(* IEC 61131-3 sources: plc-st-coding-agent/progress/evidence/f14_v12_self_20261113/jobs/diagnostic_deepseek-v4pro, 15 files *)

(* ---- public-easy-01.candidate_01.st ---- *)
(* ENGINEERING_CONTRACT
Outputs by state (state is persistent across scans):
- Pump_Motor: ON in CLEANING; starts when bottleSensor TRUE from IDLE; OFF on cleaningConfirmButton. Retained while CLEANING, even if bottleSensor falls (PUB001/PUB002).
- Filling_Valve: ON in FILLING; starts on cleaningConfirmButton in CLEANING; OFF on fillingConfirmButton (PUB002/PUB003).
- Capping_Machine: ON in CAPPING; starts on fillingConfirmButton in FILLING; OFF on cappingConfirmButton (PUB003/PUB004).
- Packing_Machine: ON in PACKING; starts on cappingConfirmButton in CAPPING; OFF on packingConfirmButton (PUB004/PUB005).
- Completion_Light: ON in COMPLETE; starts on packingConfirmButton in PACKING; reset by finishedButton (PUB005/PUB006/PUB007).
Same-scan priority: one state transition per call via ELSIF chain; outputs are assigned after transition using final state.
Buttons are treated as level-sensitive; pulse width/protocol unspecified.
*)
(* CONTRACT_RULES [] *)

FUNCTION_BLOCK FillingLineControl
VAR_INPUT
    bottleSensor: BOOL;
    cleaningConfirmButton: BOOL;
    fillingConfirmButton: BOOL;
    cappingConfirmButton: BOOL;
    packingConfirmButton: BOOL;
    finishedButton: BOOL;
END_VAR
VAR_OUTPUT
    Pump_Motor: BOOL;
    Filling_Valve: BOOL;
    Capping_Machine: BOOL;
    Packing_Machine: BOOL;
    Completion_Light: BOOL;
END_VAR
VAR
    step: INT := 0; (* 0=IDLE, 1=CLEANING, 2=FILLING, 3=CAPPING, 4=PACKING, 5=COMPLETE *)
    bottleTrig: R_TRIG;
END_VAR

(* State transitions: at most one per scan *)
bottleTrig(CLK := bottleSensor);

IF step = 0 THEN
    IF bottleTrig.Q THEN
        step := 1;
    END_IF;
ELSIF step = 1 THEN
    IF cleaningConfirmButton THEN
        step := 2;
    END_IF;
ELSIF step = 2 THEN
    IF fillingConfirmButton THEN
        step := 3;
    END_IF;
ELSIF step = 3 THEN
    IF cappingConfirmButton THEN
        step := 4;
    END_IF;
ELSIF step = 4 THEN
    IF packingConfirmButton THEN
        step := 5;
    END_IF;
ELSIF step = 5 THEN
    IF finishedButton THEN
        step := 0;
    END_IF;
END_IF;

(* Output mapping based on final state *)
CASE step OF
    0:
        Pump_Motor := FALSE;
        Filling_Valve := FALSE;
        Capping_Machine := FALSE;
        Packing_Machine := FALSE;
        Completion_Light := FALSE;

    1:
        Pump_Motor := TRUE;
        Filling_Valve := FALSE;
        Capping_Machine := FALSE;
        Packing_Machine := FALSE;
        Completion_Light := FALSE;

    2:
        Pump_Motor := FALSE;
        Filling_Valve := TRUE;
        Capping_Machine := FALSE;
        Packing_Machine := FALSE;
        Completion_Light := FALSE;

    3:
        Pump_Motor := FALSE;
        Filling_Valve := FALSE;
        Capping_Machine := TRUE;
        Packing_Machine := FALSE;
        Completion_Light := FALSE;

    4:
        Pump_Motor := FALSE;
        Filling_Valve := FALSE;
        Capping_Machine := FALSE;
        Packing_Machine := TRUE;
        Completion_Light := FALSE;

    5:
        Pump_Motor := FALSE;
        Filling_Valve := FALSE;
        Capping_Machine := FALSE;
        Packing_Machine := FALSE;
        Completion_Light := TRUE;

    ELSE
        Pump_Motor := FALSE;
        Filling_Valve := FALSE;
        Capping_Machine := FALSE;
        Packing_Machine := FALSE;
        Completion_Light := FALSE;
END_CASE;

END_FUNCTION_BLOCK

(* ---- public-easy-01.candidate_02.st ---- *)
(* ENGINEERING_CONTRACT
Outputs by state (state is persistent across scans):
- Pump_Motor: ON in CLEANING; starts when bottleSensor TRUE from IDLE; OFF on cleaningConfirmButton. Retained while CLEANING, even if bottleSensor falls (PUB001/PUB002).
- Filling_Valve: ON in FILLING; starts on cleaningConfirmButton in CLEANING; OFF on fillingConfirmButton (PUB002/PUB003).
- Capping_Machine: ON in CAPPING; starts on fillingConfirmButton in FILLING; OFF on cappingConfirmButton (PUB003/PUB004).
- Packing_Machine: ON in PACKING; starts on cappingConfirmButton in CAPPING; OFF on packingConfirmButton (PUB004/PUB005).
- Completion_Light: ON in COMPLETE; starts on packingConfirmButton in PACKING; reset by finishedButton (PUB005/PUB006/PUB007).
Same-scan priority: one state transition per call via ELSIF chain; outputs are assigned after transition using final state.
Buttons are treated as level-sensitive; pulse width/protocol unspecified.
*)
(* CONTRACT_RULES [] *)

FUNCTION_BLOCK FillingLineControl
VAR_INPUT
    bottleSensor: BOOL;
    cleaningConfirmButton: BOOL;
    fillingConfirmButton: BOOL;
    cappingConfirmButton: BOOL;
    packingConfirmButton: BOOL;
    finishedButton: BOOL;
END_VAR
VAR_OUTPUT
    Pump_Motor: BOOL;
    Filling_Valve: BOOL;
    Capping_Machine: BOOL;
    Packing_Machine: BOOL;
    Completion_Light: BOOL;
END_VAR
VAR
    step: INT := 0; (* 0=IDLE, 1=CLEANING, 2=FILLING, 3=CAPPING, 4=PACKING, 5=COMPLETE *)
END_VAR

(* State transitions: at most one per scan *)
IF step = 0 THEN
    IF bottleSensor THEN
        step := 1;
    END_IF;
ELSIF step = 1 THEN
    IF cleaningConfirmButton THEN
        step := 2;
    END_IF;
ELSIF step = 2 THEN
    IF fillingConfirmButton THEN
        step := 3;
    END_IF;
ELSIF step = 3 THEN
    IF cappingConfirmButton THEN
        step := 4;
    END_IF;
ELSIF step = 4 THEN
    IF packingConfirmButton THEN
        step := 5;
    END_IF;
ELSIF step = 5 THEN
    IF finishedButton THEN
        step := 0;
    END_IF;
END_IF;

(* Output mapping based on final state *)
CASE step OF
    0:
        Pump_Motor := FALSE;
        Filling_Valve := FALSE;
        Capping_Machine := FALSE;
        Packing_Machine := FALSE;
        Completion_Light := FALSE;

    1:
        Pump_Motor := TRUE;
        Filling_Valve := FALSE;
        Capping_Machine := FALSE;
        Packing_Machine := FALSE;
        Completion_Light := FALSE;

    2:
        Pump_Motor := FALSE;
        Filling_Valve := TRUE;
        Capping_Machine := FALSE;
        Packing_Machine := FALSE;
        Completion_Light := FALSE;

    3:
        Pump_Motor := FALSE;
        Filling_Valve := FALSE;
        Capping_Machine := TRUE;
        Packing_Machine := FALSE;
        Completion_Light := FALSE;

    4:
        Pump_Motor := FALSE;
        Filling_Valve := FALSE;
        Capping_Machine := FALSE;
        Packing_Machine := TRUE;
        Completion_Light := FALSE;

    5:
        Pump_Motor := FALSE;
        Filling_Valve := FALSE;
        Capping_Machine := FALSE;
        Packing_Machine := FALSE;
        Completion_Light := TRUE;

    ELSE
        Pump_Motor := FALSE;
        Filling_Valve := FALSE;
        Capping_Machine := FALSE;
        Packing_Machine := FALSE;
        Completion_Light := FALSE;
END_CASE;

END_FUNCTION_BLOCK

(* ---- public-easy-01.candidate_03.st ---- *)
(* ENGINEERING_CONTRACT
Outputs by state (state is persistent across scans):
- Pump_Motor: ON in CLEANING; starts when bottleSensor TRUE from IDLE; OFF on cleaningConfirmButton. Retained while CLEANING, even if bottleSensor falls (PUB001/PUB002).
- Filling_Valve: ON in FILLING; starts on cleaningConfirmButton in CLEANING; OFF on fillingConfirmButton (PUB002/PUB003).
- Capping_Machine: ON in CAPPING; starts on fillingConfirmButton in FILLING; OFF on cappingConfirmButton (PUB003/PUB004).
- Packing_Machine: ON in PACKING; starts on cappingConfirmButton in CAPPING; OFF on packingConfirmButton (PUB004/PUB005).
- Completion_Light: ON in COMPLETE; starts on packingConfirmButton in PACKING; reset by finishedButton (PUB005/PUB006/PUB007).
Same-scan priority: one state transition per call via ELSIF chain; outputs are assigned after transition using final state.
Buttons are treated as level-sensitive; pulse width/protocol unspecified.
*)
(* CONTRACT_RULES [] *)

FUNCTION_BLOCK FillingLineControl
VAR_INPUT
    bottleSensor: BOOL;
    cleaningConfirmButton: BOOL;
    fillingConfirmButton: BOOL;
    cappingConfirmButton: BOOL;
    packingConfirmButton: BOOL;
    finishedButton: BOOL;
END_VAR
VAR_OUTPUT
    Pump_Motor: BOOL;
    Filling_Valve: BOOL;
    Capping_Machine: BOOL;
    Packing_Machine: BOOL;
    Completion_Light: BOOL;
END_VAR
VAR
    step: INT := 0; (* 0=IDLE, 1=CLEANING, 2=FILLING, 3=CAPPING, 4=PACKING, 5=COMPLETE *)
    local_i: INT;
END_VAR

(* State transitions: at most one per scan *)
FOR local_i := 0 TO 5 DO
    IF step = 0 THEN
        IF bottleSensor THEN
            step := 1;
        END_IF;
    ELSIF step = 1 THEN
        IF cleaningConfirmButton THEN
            step := 2;
        END_IF;
    ELSIF step = 2 THEN
        IF fillingConfirmButton THEN
            step := 3;
        END_IF;
    ELSIF step = 3 THEN
        IF cappingConfirmButton THEN
            step := 4;
        END_IF;
    ELSIF step = 4 THEN
        IF packingConfirmButton THEN
            step := 5;
        END_IF;
    ELSIF step = 5 THEN
        IF finishedButton THEN
            step := 0;
        END_IF;
    END_IF;
END_FOR;

(* Output mapping based on final state *)
CASE step OF
    0:
        Pump_Motor := FALSE;
        Filling_Valve := FALSE;
        Capping_Machine := FALSE;
        Packing_Machine := FALSE;
        Completion_Light := FALSE;

    1:
        Pump_Motor := TRUE;
        Filling_Valve := FALSE;
        Capping_Machine := FALSE;
        Packing_Machine := FALSE;
        Completion_Light := FALSE;

    2:
        Pump_Motor := FALSE;
        Filling_Valve := TRUE;
        Capping_Machine := FALSE;
        Packing_Machine := FALSE;
        Completion_Light := FALSE;

    3:
        Pump_Motor := FALSE;
        Filling_Valve := FALSE;
        Capping_Machine := TRUE;
        Packing_Machine := FALSE;
        Completion_Light := FALSE;

    4:
        Pump_Motor := FALSE;
        Filling_Valve := FALSE;
        Capping_Machine := FALSE;
        Packing_Machine := TRUE;
        Completion_Light := FALSE;

    5:
        Pump_Motor := FALSE;
        Filling_Valve := FALSE;
        Capping_Machine := FALSE;
        Packing_Machine := FALSE;
        Completion_Light := TRUE;

    ELSE
        Pump_Motor := FALSE;
        Filling_Valve := FALSE;
        Capping_Machine := FALSE;
        Packing_Machine := FALSE;
        Completion_Light := FALSE;
END_CASE;

END_FUNCTION_BLOCK

(* ---- public-easy-01.patch_base_01.st ---- *)
(* ENGINEERING_CONTRACT
Outputs by state (state is persistent across scans):
- Pump_Motor: ON in CLEANING; starts when bottleSensor TRUE from IDLE; OFF on cleaningConfirmButton. Retained while CLEANING, even if bottleSensor falls (PUB001/PUB002).
- Filling_Valve: ON in FILLING; starts on cleaningConfirmButton in CLEANING; OFF on fillingConfirmButton (PUB002/PUB003).
- Capping_Machine: ON in CAPPING; starts on fillingConfirmButton in FILLING; OFF on cappingConfirmButton (PUB003/PUB004).
- Packing_Machine: ON in PACKING; starts on cappingConfirmButton in CAPPING; OFF on packingConfirmButton (PUB004/PUB005).
- Completion_Light: ON in COMPLETE; starts on packingConfirmButton in PACKING; reset by finishedButton (PUB005/PUB006/PUB007).
Same-scan priority: one state transition per call via ELSIF chain; outputs are assigned after transition using final state.
Buttons are treated as level-sensitive; pulse width/protocol unspecified.
*)
(* CONTRACT_RULES [] *)

FUNCTION_BLOCK FillingLineControl
VAR_INPUT
    bottleSensor: BOOL;
    cleaningConfirmButton: BOOL;
    fillingConfirmButton: BOOL;
    cappingConfirmButton: BOOL;
    packingConfirmButton: BOOL;
    finishedButton: BOOL;
END_VAR
VAR_OUTPUT
    Pump_Motor: BOOL;
    Filling_Valve: BOOL;
    Capping_Machine: BOOL;
    Packing_Machine: BOOL;
    Completion_Light: BOOL;
END_VAR
VAR
    step: INT := 0; (* 0=IDLE, 1=CLEANING, 2=FILLING, 3=CAPPING, 4=PACKING, 5=COMPLETE *)
END_VAR

(* State transitions: at most one per scan *)
IF step = 0 THEN
    IF bottleSensor THEN
        step := 1;
    END_IF;
ELSIF step = 1 THEN
    IF cleaningConfirmButton THEN
        step := 2;
    END_IF;
ELSIF step = 2 THEN
    IF fillingConfirmButton THEN
        step := 3;
    END_IF;
ELSIF step = 3 THEN
    IF cappingConfirmButton THEN
        step := 4;
    END_IF;
ELSIF step = 4 THEN
    IF packingConfirmButton THEN
        step := 5;
    END_IF;
ELSIF step = 5 THEN
    IF finishedButton THEN
        step := 0;
    END_IF;
END_IF;

(* Output mapping based on final state *)
CASE step OF
    0:
        Pump_Motor := FALSE;
        Filling_Valve := FALSE;
        Capping_Machine := FALSE;
        Packing_Machine := FALSE;
        Completion_Light := FALSE;

    1:
        Pump_Motor := TRUE;
        Filling_Valve := FALSE;
        Capping_Machine := FALSE;
        Packing_Machine := FALSE;
        Completion_Light := FALSE;

    2:
        Pump_Motor := FALSE;
        Filling_Valve := TRUE;
        Capping_Machine := FALSE;
        Packing_Machine := FALSE;
        Completion_Light := FALSE;

    3:
        Pump_Motor := FALSE;
        Filling_Valve := FALSE;
        Capping_Machine := TRUE;
        Packing_Machine := FALSE;
        Completion_Light := FALSE;

    4:
        Pump_Motor := FALSE;
        Filling_Valve := FALSE;
        Capping_Machine := FALSE;
        Packing_Machine := TRUE;
        Completion_Light := FALSE;

    5:
        Pump_Motor := FALSE;
        Filling_Valve := FALSE;
        Capping_Machine := FALSE;
        Packing_Machine := FALSE;
        Completion_Light := TRUE;

    ELSE
        Pump_Motor := FALSE;
        Filling_Valve := FALSE;
        Capping_Machine := FALSE;
        Packing_Machine := FALSE;
        Completion_Light := FALSE;
END_CASE;

END_FUNCTION_BLOCK

(* ---- public-easy-01.patch_base_02.st ---- *)
(* ENGINEERING_CONTRACT
Outputs by state (state is persistent across scans):
- Pump_Motor: ON in CLEANING; starts when bottleSensor TRUE from IDLE; OFF on cleaningConfirmButton. Retained while CLEANING, even if bottleSensor falls (PUB001/PUB002).
- Filling_Valve: ON in FILLING; starts on cleaningConfirmButton in CLEANING; OFF on fillingConfirmButton (PUB002/PUB003).
- Capping_Machine: ON in CAPPING; starts on fillingConfirmButton in FILLING; OFF on cappingConfirmButton (PUB003/PUB004).
- Packing_Machine: ON in PACKING; starts on cappingConfirmButton in CAPPING; OFF on packingConfirmButton (PUB004/PUB005).
- Completion_Light: ON in COMPLETE; starts on packingConfirmButton in PACKING; reset by finishedButton (PUB005/PUB006/PUB007).
Same-scan priority: one state transition per call via ELSIF chain; outputs are assigned after transition using final state.
Buttons are treated as level-sensitive; pulse width/protocol unspecified.
*)
(* CONTRACT_RULES [] *)

FUNCTION_BLOCK FillingLineControl
VAR_INPUT
    bottleSensor: BOOL;
    cleaningConfirmButton: BOOL;
    fillingConfirmButton: BOOL;
    cappingConfirmButton: BOOL;
    packingConfirmButton: BOOL;
    finishedButton: BOOL;
END_VAR
VAR_OUTPUT
    Pump_Motor: BOOL;
    Filling_Valve: BOOL;
    Capping_Machine: BOOL;
    Packing_Machine: BOOL;
    Completion_Light: BOOL;
END_VAR
VAR
    step: INT := 0; (* 0=IDLE, 1=CLEANING, 2=FILLING, 3=CAPPING, 4=PACKING, 5=COMPLETE *)
    bottleTrig: R_TRIG;
END_VAR

(* State transitions: at most one per scan *)
bottleTrig(CLK := bottleSensor);

IF step = 0 THEN
    IF bottleTrig.Q THEN
        step := 1;
    END_IF;
ELSIF step = 1 THEN
    IF cleaningConfirmButton THEN
        step := 2;
    END_IF;
ELSIF step = 2 THEN
    IF fillingConfirmButton THEN
        step := 3;
    END_IF;
ELSIF step = 3 THEN
    IF cappingConfirmButton THEN
        step := 4;
    END_IF;
ELSIF step = 4 THEN
    IF packingConfirmButton THEN
        step := 5;
    END_IF;
ELSIF step = 5 THEN
    IF finishedButton THEN
        step := 0;
    END_IF;
END_IF;

(* Output mapping based on final state *)
CASE step OF
    0:
        Pump_Motor := FALSE;
        Filling_Valve := FALSE;
        Capping_Machine := FALSE;
        Packing_Machine := FALSE;
        Completion_Light := FALSE;

    1:
        Pump_Motor := TRUE;
        Filling_Valve := FALSE;
        Capping_Machine := FALSE;
        Packing_Machine := FALSE;
        Completion_Light := FALSE;

    2:
        Pump_Motor := FALSE;
        Filling_Valve := TRUE;
        Capping_Machine := FALSE;
        Packing_Machine := FALSE;
        Completion_Light := FALSE;

    3:
        Pump_Motor := FALSE;
        Filling_Valve := FALSE;
        Capping_Machine := TRUE;
        Packing_Machine := FALSE;
        Completion_Light := FALSE;

    4:
        Pump_Motor := FALSE;
        Filling_Valve := FALSE;
        Capping_Machine := FALSE;
        Packing_Machine := TRUE;
        Completion_Light := FALSE;

    5:
        Pump_Motor := FALSE;
        Filling_Valve := FALSE;
        Capping_Machine := FALSE;
        Packing_Machine := FALSE;
        Completion_Light := TRUE;

    ELSE
        Pump_Motor := FALSE;
        Filling_Valve := FALSE;
        Capping_Machine := FALSE;
        Packing_Machine := FALSE;
        Completion_Light := FALSE;
END_CASE;

END_FUNCTION_BLOCK

(* ---- public-easy-01.patch_base_03.st ---- *)
(* ENGINEERING_CONTRACT
Outputs by state (state is persistent across scans):
- Pump_Motor: ON in CLEANING; starts when bottleSensor TRUE from IDLE; OFF on cleaningConfirmButton. Retained while CLEANING, even if bottleSensor falls (PUB001/PUB002).
- Filling_Valve: ON in FILLING; starts on cleaningConfirmButton in CLEANING; OFF on fillingConfirmButton (PUB002/PUB003).
- Capping_Machine: ON in CAPPING; starts on fillingConfirmButton in FILLING; OFF on cappingConfirmButton (PUB003/PUB004).
- Packing_Machine: ON in PACKING; starts on cappingConfirmButton in CAPPING; OFF on packingConfirmButton (PUB004/PUB005).
- Completion_Light: ON in COMPLETE; starts on packingConfirmButton in PACKING; reset by finishedButton (PUB005/PUB006/PUB007).
Same-scan priority: one state transition per call via ELSIF chain; outputs are assigned after transition using final state.
Buttons are treated as level-sensitive; pulse width/protocol unspecified.
*)
(* CONTRACT_RULES [] *)

FUNCTION_BLOCK FillingLineControl
VAR_INPUT
    bottleSensor: BOOL;
    cleaningConfirmButton: BOOL;
    fillingConfirmButton: BOOL;
    cappingConfirmButton: BOOL;
    packingConfirmButton: BOOL;
    finishedButton: BOOL;
END_VAR
VAR_OUTPUT
    Pump_Motor: BOOL;
    Filling_Valve: BOOL;
    Capping_Machine: BOOL;
    Packing_Machine: BOOL;
    Completion_Light: BOOL;
END_VAR
VAR
    step: INT := 0; (* 0=IDLE, 1=CLEANING, 2=FILLING, 3=CAPPING, 4=PACKING, 5=COMPLETE *)
END_VAR

(* State transitions: at most one per scan *)
IF step = 0 THEN
    IF bottleSensor THEN
        step := 1;
    END_IF;
ELSIF step = 1 THEN
    IF cleaningConfirmButton THEN
        step := 2;
    END_IF;
ELSIF step = 2 THEN
    IF fillingConfirmButton THEN
        step := 3;
    END_IF;
ELSIF step = 3 THEN
    IF cappingConfirmButton THEN
        step := 4;
    END_IF;
ELSIF step = 4 THEN
    IF packingConfirmButton THEN
        step := 5;
    END_IF;
ELSIF step = 5 THEN
    IF finishedButton THEN
        step := 0;
    END_IF;
END_IF;

(* Output mapping based on final state *)
CASE step OF
    0:
        Pump_Motor := FALSE;
        Filling_Valve := FALSE;
        Capping_Machine := FALSE;
        Packing_Machine := FALSE;
        Completion_Light := FALSE;

    1:
        Pump_Motor := TRUE;
        Filling_Valve := FALSE;
        Capping_Machine := FALSE;
        Packing_Machine := FALSE;
        Completion_Light := FALSE;

    2:
        Pump_Motor := FALSE;
        Filling_Valve := TRUE;
        Capping_Machine := FALSE;
        Packing_Machine := FALSE;
        Completion_Light := FALSE;

    3:
        Pump_Motor := FALSE;
        Filling_Valve := FALSE;
        Capping_Machine := TRUE;
        Packing_Machine := FALSE;
        Completion_Light := FALSE;

    4:
        Pump_Motor := FALSE;
        Filling_Valve := FALSE;
        Capping_Machine := FALSE;
        Packing_Machine := TRUE;
        Completion_Light := FALSE;

    5:
        Pump_Motor := FALSE;
        Filling_Valve := FALSE;
        Capping_Machine := FALSE;
        Packing_Machine := FALSE;
        Completion_Light := TRUE;

    ELSE
        Pump_Motor := FALSE;
        Filling_Valve := FALSE;
        Capping_Machine := FALSE;
        Packing_Machine := FALSE;
        Completion_Light := FALSE;
END_CASE;

END_FUNCTION_BLOCK

(* ---- public-easy-01.raw_candidate_01.st ---- *)
(* ENGINEERING_CONTRACT
Outputs by state (state is persistent across scans):
- Pump_Motor: ON in CLEANING; starts when bottleSensor TRUE from IDLE; OFF on cleaningConfirmButton. Retained while CLEANING, even if bottleSensor falls (PUB001/PUB002).
- Filling_Valve: ON in FILLING; starts on cleaningConfirmButton in CLEANING; OFF on fillingConfirmButton (PUB002/PUB003).
- Capping_Machine: ON in CAPPING; starts on fillingConfirmButton in FILLING; OFF on cappingConfirmButton (PUB003/PUB004).
- Packing_Machine: ON in PACKING; starts on cappingConfirmButton in CAPPING; OFF on packingConfirmButton (PUB004/PUB005).
- Completion_Light: ON in COMPLETE; starts on packingConfirmButton in PACKING; reset by finishedButton (PUB005/PUB006/PUB007).
Same-scan priority: one state transition per call via ELSIF chain; outputs are assigned after transition using final state.
Buttons are treated as level-sensitive; pulse width/protocol unspecified.
*)
(* CONTRACT_RULES [] *)

FUNCTION_BLOCK FillingLineControl
VAR_INPUT
    bottleSensor: BOOL;
    cleaningConfirmButton: BOOL;
    fillingConfirmButton: BOOL;
    cappingConfirmButton: BOOL;
    packingConfirmButton: BOOL;
    finishedButton: BOOL;
END_VAR
VAR_OUTPUT
    Pump_Motor: BOOL;
    Filling_Valve: BOOL;
    Capping_Machine: BOOL;
    Packing_Machine: BOOL;
    Completion_Light: BOOL;
END_VAR
VAR
    step: INT := 0; (* 0=IDLE, 1=CLEANING, 2=FILLING, 3=CAPPING, 4=PACKING, 5=COMPLETE *)
    bottleTrig: R_TRIG;
END_VAR

(* State transitions: at most one per scan *)
bottleTrig(CLK := bottleSensor);

IF step = 0 THEN
    IF bottleTrig.Q THEN
        step := 1;
    END_IF;
ELSIF step = 1 THEN
    IF cleaningConfirmButton THEN
        step := 2;
    END_IF;
ELSIF step = 2 THEN
    IF fillingConfirmButton THEN
        step := 3;
    END_IF;
ELSIF step = 3 THEN
    IF cappingConfirmButton THEN
        step := 4;
    END_IF;
ELSIF step = 4 THEN
    IF packingConfirmButton THEN
        step := 5;
    END_IF;
ELSIF step = 5 THEN
    IF finishedButton THEN
        step := 0;
    END_IF;
END_IF;

(* Output mapping based on final state *)
CASE step OF
    0:
        Pump_Motor := FALSE;
        Filling_Valve := FALSE;
        Capping_Machine := FALSE;
        Packing_Machine := FALSE;
        Completion_Light := FALSE;

    1:
        Pump_Motor := TRUE;
        Filling_Valve := FALSE;
        Capping_Machine := FALSE;
        Packing_Machine := FALSE;
        Completion_Light := FALSE;

    2:
        Pump_Motor := FALSE;
        Filling_Valve := TRUE;
        Capping_Machine := FALSE;
        Packing_Machine := FALSE;
        Completion_Light := FALSE;

    3:
        Pump_Motor := FALSE;
        Filling_Valve := FALSE;
        Capping_Machine := TRUE;
        Packing_Machine := FALSE;
        Completion_Light := FALSE;

    4:
        Pump_Motor := FALSE;
        Filling_Valve := FALSE;
        Capping_Machine := FALSE;
        Packing_Machine := TRUE;
        Completion_Light := FALSE;

    5:
        Pump_Motor := FALSE;
        Filling_Valve := FALSE;
        Capping_Machine := FALSE;
        Packing_Machine := FALSE;
        Completion_Light := TRUE;

    ELSE
        Pump_Motor := FALSE;
        Filling_Valve := FALSE;
        Capping_Machine := FALSE;
        Packing_Machine := FALSE;
        Completion_Light := FALSE;
END_CASE;

END_FUNCTION_BLOCK

(* ---- public-easy-01.raw_candidate_02.st ---- *)
(* ENGINEERING_CONTRACT
Outputs by state (state is persistent across scans):
- Pump_Motor: ON in CLEANING; starts when bottleSensor TRUE from IDLE; OFF on cleaningConfirmButton. Retained while CLEANING, even if bottleSensor falls (PUB001/PUB002).
- Filling_Valve: ON in FILLING; starts on cleaningConfirmButton in CLEANING; OFF on fillingConfirmButton (PUB002/PUB003).
- Capping_Machine: ON in CAPPING; starts on fillingConfirmButton in FILLING; OFF on cappingConfirmButton (PUB003/PUB004).
- Packing_Machine: ON in PACKING; starts on cappingConfirmButton in CAPPING; OFF on packingConfirmButton (PUB004/PUB005).
- Completion_Light: ON in COMPLETE; starts on packingConfirmButton in PACKING; reset by finishedButton (PUB005/PUB006/PUB007).
Same-scan priority: one state transition per call via ELSIF chain; outputs are assigned after transition using final state.
Buttons are treated as level-sensitive; pulse width/protocol unspecified.
*)
(* CONTRACT_RULES [] *)

FUNCTION_BLOCK FillingLineControl
VAR_INPUT
    bottleSensor: BOOL;
    cleaningConfirmButton: BOOL;
    fillingConfirmButton: BOOL;
    cappingConfirmButton: BOOL;
    packingConfirmButton: BOOL;
    finishedButton: BOOL;
END_VAR
VAR_OUTPUT
    Pump_Motor: BOOL;
    Filling_Valve: BOOL;
    Capping_Machine: BOOL;
    Packing_Machine: BOOL;
    Completion_Light: BOOL;
END_VAR
VAR
    step: INT := 0; (* 0=IDLE, 1=CLEANING, 2=FILLING, 3=CAPPING, 4=PACKING, 5=COMPLETE *)
END_VAR

(* State transitions: at most one per scan *)
IF step = 0 THEN
    IF bottleSensor THEN
        step := 1;
    END_IF;
ELSIF step = 1 THEN
    IF cleaningConfirmButton THEN
        step := 2;
    END_IF;
ELSIF step = 2 THEN
    IF fillingConfirmButton THEN
        step := 3;
    END_IF;
ELSIF step = 3 THEN
    IF cappingConfirmButton THEN
        step := 4;
    END_IF;
ELSIF step = 4 THEN
    IF packingConfirmButton THEN
        step := 5;
    END_IF;
ELSIF step = 5 THEN
    IF finishedButton THEN
        step := 0;
    END_IF;
END_IF;

(* Output mapping based on final state *)
CASE step OF
    0:
        Pump_Motor := FALSE;
        Filling_Valve := FALSE;
        Capping_Machine := FALSE;
        Packing_Machine := FALSE;
        Completion_Light := FALSE;

    1:
        Pump_Motor := TRUE;
        Filling_Valve := FALSE;
        Capping_Machine := FALSE;
        Packing_Machine := FALSE;
        Completion_Light := FALSE;

    2:
        Pump_Motor := FALSE;
        Filling_Valve := TRUE;
        Capping_Machine := FALSE;
        Packing_Machine := FALSE;
        Completion_Light := FALSE;

    3:
        Pump_Motor := FALSE;
        Filling_Valve := FALSE;
        Capping_Machine := TRUE;
        Packing_Machine := FALSE;
        Completion_Light := FALSE;

    4:
        Pump_Motor := FALSE;
        Filling_Valve := FALSE;
        Capping_Machine := FALSE;
        Packing_Machine := TRUE;
        Completion_Light := FALSE;

    5:
        Pump_Motor := FALSE;
        Filling_Valve := FALSE;
        Capping_Machine := FALSE;
        Packing_Machine := FALSE;
        Completion_Light := TRUE;

    ELSE
        Pump_Motor := FALSE;
        Filling_Valve := FALSE;
        Capping_Machine := FALSE;
        Packing_Machine := FALSE;
        Completion_Light := FALSE;
END_CASE;

END_FUNCTION_BLOCK

(* ---- public-easy-01.raw_candidate_03.st ---- *)
(* ENGINEERING_CONTRACT
Outputs by state (state is persistent across scans):
- Pump_Motor: ON in CLEANING; starts when bottleSensor TRUE from IDLE; OFF on cleaningConfirmButton. Retained while CLEANING, even if bottleSensor falls (PUB001/PUB002).
- Filling_Valve: ON in FILLING; starts on cleaningConfirmButton in CLEANING; OFF on fillingConfirmButton (PUB002/PUB003).
- Capping_Machine: ON in CAPPING; starts on fillingConfirmButton in FILLING; OFF on cappingConfirmButton (PUB003/PUB004).
- Packing_Machine: ON in PACKING; starts on cappingConfirmButton in CAPPING; OFF on packingConfirmButton (PUB004/PUB005).
- Completion_Light: ON in COMPLETE; starts on packingConfirmButton in PACKING; reset by finishedButton (PUB005/PUB006/PUB007).
Same-scan priority: one state transition per call via ELSIF chain; outputs are assigned after transition using final state.
Buttons are treated as level-sensitive; pulse width/protocol unspecified.
*)
(* CONTRACT_RULES [] *)

FUNCTION_BLOCK FillingLineControl
VAR_INPUT
    bottleSensor: BOOL;
    cleaningConfirmButton: BOOL;
    fillingConfirmButton: BOOL;
    cappingConfirmButton: BOOL;
    packingConfirmButton: BOOL;
    finishedButton: BOOL;
END_VAR
VAR_OUTPUT
    Pump_Motor: BOOL;
    Filling_Valve: BOOL;
    Capping_Machine: BOOL;
    Packing_Machine: BOOL;
    Completion_Light: BOOL;
END_VAR
VAR
    step: INT := 0; (* 0=IDLE, 1=CLEANING, 2=FILLING, 3=CAPPING, 4=PACKING, 5=COMPLETE *)
    local_i: INT;
END_VAR

(* State transitions: at most one per scan *)
FOR local_i := 0 TO 5 DO
    IF step = 0 THEN
        IF bottleSensor THEN
            step := 1;
        END_IF;
    ELSIF step = 1 THEN
        IF cleaningConfirmButton THEN
            step := 2;
        END_IF;
    ELSIF step = 2 THEN
        IF fillingConfirmButton THEN
            step := 3;
        END_IF;
    ELSIF step = 3 THEN
        IF cappingConfirmButton THEN
            step := 4;
        END_IF;
    ELSIF step = 4 THEN
        IF packingConfirmButton THEN
            step := 5;
        END_IF;
    ELSIF step = 5 THEN
        IF finishedButton THEN
            step := 0;
        END_IF;
    END_IF;
END_FOR;

(* Output mapping based on final state *)
CASE step OF
    0:
        Pump_Motor := FALSE;
        Filling_Valve := FALSE;
        Capping_Machine := FALSE;
        Packing_Machine := FALSE;
        Completion_Light := FALSE;

    1:
        Pump_Motor := TRUE;
        Filling_Valve := FALSE;
        Capping_Machine := FALSE;
        Packing_Machine := FALSE;
        Completion_Light := FALSE;

    2:
        Pump_Motor := FALSE;
        Filling_Valve := TRUE;
        Capping_Machine := FALSE;
        Packing_Machine := FALSE;
        Completion_Light := FALSE;

    3:
        Pump_Motor := FALSE;
        Filling_Valve := FALSE;
        Capping_Machine := TRUE;
        Packing_Machine := FALSE;
        Completion_Light := FALSE;

    4:
        Pump_Motor := FALSE;
        Filling_Valve := FALSE;
        Capping_Machine := FALSE;
        Packing_Machine := TRUE;
        Completion_Light := FALSE;

    5:
        Pump_Motor := FALSE;
        Filling_Valve := FALSE;
        Capping_Machine := FALSE;
        Packing_Machine := FALSE;
        Completion_Light := TRUE;

    ELSE
        Pump_Motor := FALSE;
        Filling_Valve := FALSE;
        Capping_Machine := FALSE;
        Packing_Machine := FALSE;
        Completion_Light := FALSE;
END_CASE;

END_FUNCTION_BLOCK

(* ---- public-hard-05.candidate_01.st ---- *)
(* ENGINEERING_CONTRACT
Manual: moving/grip/release outputs are combinational from corresponding button AND NOT corresponding limit switch; releasing the button clears the output. PUB001, PUB005.
SingleStep: rising Start advances only when idle or current step limit reached; each step holds its output until its limit, then waits for next Start. After step 8, next Start goes to step 1. PUB002.
SingleCycle: rising Start starts step 1; each step auto-advances on its completion limit, then stops at step 0 after step 8. PUB003.
Continuous: rising Start starts step 1; auto-advances and loops 8->1. PUB004.
EmergencyStop=FALSE forces all outputs FALSE and freezes automatic state changes. No reset is inferred. PUB005.
Completion feedback uses DownLimitSwitch, UpLimitSwitch, LeftLimitSwitch, RightLimitSwitch, GripLimitSwitch, ReleaseLimitSwitch. Unspecified mode-change behavior preserves the automatic step state.
*)
(* CONTRACT_RULES [] *)
FUNCTION_BLOCK FB_MechanicalArmControl
VAR_INPUT
    ManualMode : BOOL;
    SingleStepMode : BOOL;
    SingleCycleMode : BOOL;
    ContinuousMode : BOOL;
    EmergencyStop : BOOL;
    Start : BOOL;
    DownButton : BOOL;
    UpButton : BOOL;
    LeftButton : BOOL;
    RightButton : BOOL;
    GripButton : BOOL;
    ReleaseButton : BOOL;
    DownLimitSwitch : BOOL;
    UpLimitSwitch : BOOL;
    LeftLimitSwitch : BOOL;
    RightLimitSwitch : BOOL;
    GripLimitSwitch : BOOL;
    ReleaseLimitSwitch : BOOL;
END_VAR
VAR_OUTPUT
    MoveDown : BOOL;
    MoveUp : BOOL;
    MoveLeft : BOOL;
    MoveRight : BOOL;
    ActivateGrip : BOOL;
    ActivateRelease : BOOL;
END_VAR
VAR
    startTrig : R_TRIG;
    sdStep : INT := 0;
    autoStep : INT := 0;
    sdDone : BOOL;
    autoDone : BOOL;
    tmpMoveDown : BOOL;
    tmpMoveUp : BOOL;
    tmpMoveLeft : BOOL;
    tmpMoveRight : BOOL;
    tmpActivateGrip : BOOL;
    tmpActivateRelease : BOOL;
END_VAR

startTrig(CLK := Start);

tmpMoveDown := FALSE;
tmpMoveUp := FALSE;
tmpMoveLeft := FALSE;
tmpMoveRight := FALSE;
tmpActivateGrip := FALSE;
tmpActivateRelease := FALSE;

IF ManualMode THEN
    tmpMoveDown := DownButton AND NOT DownLimitSwitch;
    tmpMoveUp := UpButton AND NOT UpLimitSwitch;
    tmpMoveLeft := LeftButton AND NOT LeftLimitSwitch;
    tmpMoveRight := RightButton AND NOT RightLimitSwitch;
    tmpActivateGrip := GripButton AND NOT GripLimitSwitch;
    tmpActivateRelease := ReleaseButton AND NOT ReleaseLimitSwitch;

    IF tmpMoveDown AND tmpMoveUp THEN
        tmpMoveDown := FALSE;
        tmpMoveUp := FALSE;
    END_IF;
    IF tmpMoveLeft AND tmpMoveRight THEN
        tmpMoveLeft := FALSE;
        tmpMoveRight := FALSE;
    END_IF;
    IF tmpActivateGrip AND tmpActivateRelease THEN
        tmpActivateGrip := FALSE;
        tmpActivateRelease := FALSE;
    END_IF;

ELSIF SingleStepMode THEN
    CASE sdStep OF
        1: sdDone := DownLimitSwitch;
        2: sdDone := GripLimitSwitch;
        3: sdDone := UpLimitSwitch;
        4: sdDone := RightLimitSwitch;
        5: sdDone := DownLimitSwitch;
        6: sdDone := ReleaseLimitSwitch;
        7: sdDone := UpLimitSwitch;
        8: sdDone := LeftLimitSwitch;
    ELSE
        sdDone := TRUE;
    END_CASE;

    IF EmergencyStop AND startTrig.Q AND sdDone THEN
        IF sdStep >= 8 THEN
            sdStep := 1;
        ELSE
            sdStep := sdStep + 1;
        END_IF;
    END_IF;

    CASE sdStep OF
        1: tmpMoveDown := NOT DownLimitSwitch;
        2: tmpActivateGrip := NOT GripLimitSwitch;
        3: tmpMoveUp := NOT UpLimitSwitch;
        4: tmpMoveRight := NOT RightLimitSwitch;
        5: tmpMoveDown := NOT DownLimitSwitch;
        6: tmpActivateRelease := NOT ReleaseLimitSwitch;
        7: tmpMoveUp := NOT UpLimitSwitch;
        8: tmpMoveLeft := NOT LeftLimitSwitch;
    END_CASE;

ELSIF (SingleCycleMode OR ContinuousMode) THEN
    IF EmergencyStop AND startTrig.Q AND (autoStep = 0) THEN
        autoStep := 1;
    END_IF;

    CASE autoStep OF
        1: autoDone := DownLimitSwitch;
        2: autoDone := GripLimitSwitch;
        3: autoDone := UpLimitSwitch;
        4: autoDone := RightLimitSwitch;
        5: autoDone := DownLimitSwitch;
        6: autoDone := ReleaseLimitSwitch;
        7: autoDone := UpLimitSwitch;
        8: autoDone := LeftLimitSwitch;
    ELSE
        autoDone := TRUE;
    END_CASE;

    IF EmergencyStop AND (autoStep <> 0) AND autoDone THEN
        IF SingleCycleMode THEN
            IF autoStep < 8 THEN
                autoStep := autoStep + 1;
            ELSE
                autoStep := 0;
            END_IF;
        ELSIF ContinuousMode THEN
            IF autoStep < 8 THEN
                autoStep := autoStep + 1;
            ELSE
                autoStep := 1;
            END_IF;
        END_IF;
    END_IF;

    CASE autoStep OF
        1: tmpMoveDown := NOT DownLimitSwitch;
        2: tmpActivateGrip := NOT GripLimitSwitch;
        3: tmpMoveUp := NOT UpLimitSwitch;
        4: tmpMoveRight := NOT RightLimitSwitch;
        5: tmpMoveDown := NOT DownLimitSwitch;
        6: tmpActivateRelease := NOT ReleaseLimitSwitch;
        7: tmpMoveUp := NOT UpLimitSwitch;
        8: tmpMoveLeft := NOT LeftLimitSwitch;
    END_CASE;

END_IF;

IF NOT EmergencyStop THEN
    MoveDown := FALSE;
    MoveUp := FALSE;
    MoveLeft := FALSE;
    MoveRight := FALSE;
    ActivateGrip := FALSE;
    ActivateRelease := FALSE;
ELSE
    MoveDown := tmpMoveDown;
    MoveUp := tmpMoveUp;
    MoveLeft := tmpMoveLeft;
    MoveRight := tmpMoveRight;
    ActivateGrip := tmpActivateGrip;
    ActivateRelease := tmpActivateRelease;
END_IF;

END_FUNCTION_BLOCK

(* ---- public-hard-05.patch_base_01.st ---- *)
(* ENGINEERING_CONTRACT
Manual: moving/grip/release outputs are combinational from corresponding button AND NOT corresponding limit switch; releasing the button clears the output. PUB001, PUB005.
SingleStep: rising Start advances only when idle or current step limit reached; each step holds its output until its limit, then waits for next Start. After step 8, next Start goes to step 1. PUB002.
SingleCycle: rising Start starts step 1; each step auto-advances on its completion limit, then stops at step 0 after step 8. PUB003.
Continuous: rising Start starts step 1; auto-advances and loops 8->1. PUB004.
EmergencyStop=FALSE forces all outputs FALSE and freezes automatic state changes. No reset is inferred. PUB005.
Completion feedback uses DownLimitSwitch, UpLimitSwitch, LeftLimitSwitch, RightLimitSwitch, GripLimitSwitch, ReleaseLimitSwitch. Unspecified mode-change behavior preserves the automatic step state.
*)
(* CONTRACT_RULES [] *)
FUNCTION_BLOCK FB_MechanicalArmControl
VAR_INPUT
    ManualMode : BOOL;
    SingleStepMode : BOOL;
    SingleCycleMode : BOOL;
    ContinuousMode : BOOL;
    EmergencyStop : BOOL;
    Start : BOOL;
    DownButton : BOOL;
    UpButton : BOOL;
    LeftButton : BOOL;
    RightButton : BOOL;
    GripButton : BOOL;
    ReleaseButton : BOOL;
    DownLimitSwitch : BOOL;
    UpLimitSwitch : BOOL;
    LeftLimitSwitch : BOOL;
    RightLimitSwitch : BOOL;
    GripLimitSwitch : BOOL;
    ReleaseLimitSwitch : BOOL;
END_VAR
VAR_OUTPUT
    MoveDown : BOOL;
    MoveUp : BOOL;
    MoveLeft : BOOL;
    MoveRight : BOOL;
    ActivateGrip : BOOL;
    ActivateRelease : BOOL;
END_VAR
VAR
    startTrig : R_TRIG;
    sdStep : INT := 0;
    autoStep : INT := 0;
    sdDone : BOOL;
    autoDone : BOOL;
    tmpMoveDown : BOOL;
    tmpMoveUp : BOOL;
    tmpMoveLeft : BOOL;
    tmpMoveRight : BOOL;
    tmpActivateGrip : BOOL;
    tmpActivateRelease : BOOL;
END_VAR

startTrig(CLK := Start);

tmpMoveDown := FALSE;
tmpMoveUp := FALSE;
tmpMoveLeft := FALSE;
tmpMoveRight := FALSE;
tmpActivateGrip := FALSE;
tmpActivateRelease := FALSE;

IF ManualMode THEN
    tmpMoveDown := DownButton AND NOT DownLimitSwitch;
    tmpMoveUp := UpButton AND NOT UpLimitSwitch;
    tmpMoveLeft := LeftButton AND NOT LeftLimitSwitch;
    tmpMoveRight := RightButton AND NOT RightLimitSwitch;
    tmpActivateGrip := GripButton AND NOT GripLimitSwitch;
    tmpActivateRelease := ReleaseButton AND NOT ReleaseLimitSwitch;

ELSIF SingleStepMode THEN
    CASE sdStep OF
        1: sdDone := DownLimitSwitch;
        2: sdDone := GripLimitSwitch;
        3: sdDone := UpLimitSwitch;
        4: sdDone := RightLimitSwitch;
        5: sdDone := DownLimitSwitch;
        6: sdDone := ReleaseLimitSwitch;
        7: sdDone := UpLimitSwitch;
        8: sdDone := LeftLimitSwitch;
    ELSE
        sdDone := TRUE;
    END_CASE;

    IF EmergencyStop AND startTrig.Q AND sdDone THEN
        IF sdStep >= 8 THEN
            sdStep := 1;
        ELSE
            sdStep := sdStep + 1;
        END_IF;
    END_IF;

    CASE sdStep OF
        1: tmpMoveDown := NOT DownLimitSwitch;
        2: tmpActivateGrip := NOT GripLimitSwitch;
        3: tmpMoveUp := NOT UpLimitSwitch;
        4: tmpMoveRight := NOT RightLimitSwitch;
        5: tmpMoveDown := NOT DownLimitSwitch;
        6: tmpActivateRelease := NOT ReleaseLimitSwitch;
        7: tmpMoveUp := NOT UpLimitSwitch;
        8: tmpMoveLeft := NOT LeftLimitSwitch;
    END_CASE;

ELSIF (SingleCycleMode OR ContinuousMode) THEN
    IF EmergencyStop AND startTrig.Q AND (autoStep = 0) THEN
        autoStep := 1;
    END_IF;

    CASE autoStep OF
        1: autoDone := DownLimitSwitch;
        2: autoDone := GripLimitSwitch;
        3: autoDone := UpLimitSwitch;
        4: autoDone := RightLimitSwitch;
        5: autoDone := DownLimitSwitch;
        6: autoDone := ReleaseLimitSwitch;
        7: autoDone := UpLimitSwitch;
        8: autoDone := LeftLimitSwitch;
    ELSE
        autoDone := TRUE;
    END_CASE;

    IF EmergencyStop AND (autoStep <> 0) AND autoDone THEN
        IF SingleCycleMode THEN
            IF autoStep < 8 THEN
                autoStep := autoStep + 1;
            ELSE
                autoStep := 0;
            END_IF;
        ELSIF ContinuousMode THEN
            IF autoStep < 8 THEN
                autoStep := autoStep + 1;
            ELSE
                autoStep := 1;
            END_IF;
        END_IF;
    END_IF;

    CASE autoStep OF
        1: tmpMoveDown := NOT DownLimitSwitch;
        2: tmpActivateGrip := NOT GripLimitSwitch;
        3: tmpMoveUp := NOT UpLimitSwitch;
        4: tmpMoveRight := NOT RightLimitSwitch;
        5: tmpMoveDown := NOT DownLimitSwitch;
        6: tmpActivateRelease := NOT ReleaseLimitSwitch;
        7: tmpMoveUp := NOT UpLimitSwitch;
        8: tmpMoveLeft := NOT LeftLimitSwitch;
    END_CASE;

END_IF;

IF NOT EmergencyStop THEN
    MoveDown := FALSE;
    MoveUp := FALSE;
    MoveLeft := FALSE;
    MoveRight := FALSE;
    ActivateGrip := FALSE;
    ActivateRelease := FALSE;
ELSE
    MoveDown := tmpMoveDown;
    MoveUp := tmpMoveUp;
    MoveLeft := tmpMoveLeft;
    MoveRight := tmpMoveRight;
    ActivateGrip := tmpActivateGrip;
    ActivateRelease := tmpActivateRelease;
END_IF;

END_FUNCTION_BLOCK

(* ---- public-hard-05.raw_candidate_01.st ---- *)
(* ENGINEERING_CONTRACT
Manual: moving/grip/release outputs are combinational from corresponding button AND NOT corresponding limit switch; releasing the button clears the output. PUB001, PUB005.
SingleStep: rising Start advances only when idle or current step limit reached; each step holds its output until its limit, then waits for next Start. After step 8, next Start goes to step 1. PUB002.
SingleCycle: rising Start starts step 1; each step auto-advances on its completion limit, then stops at step 0 after step 8. PUB003.
Continuous: rising Start starts step 1; auto-advances and loops 8->1. PUB004.
EmergencyStop=FALSE forces all outputs FALSE and freezes automatic state changes. No reset is inferred. PUB005.
Completion feedback uses DownLimitSwitch, UpLimitSwitch, LeftLimitSwitch, RightLimitSwitch, GripLimitSwitch, ReleaseLimitSwitch. Unspecified mode-change behavior preserves the automatic step state.
*)
(* CONTRACT_RULES [] *)
FUNCTION_BLOCK FB_MechanicalArmControl
VAR_INPUT
    ManualMode : BOOL;
    SingleStepMode : BOOL;
    SingleCycleMode : BOOL;
    ContinuousMode : BOOL;
    EmergencyStop : BOOL;
    Start : BOOL;
    DownButton : BOOL;
    UpButton : BOOL;
    LeftButton : BOOL;
    RightButton : BOOL;
    GripButton : BOOL;
    ReleaseButton : BOOL;
    DownLimitSwitch : BOOL;
    UpLimitSwitch : BOOL;
    LeftLimitSwitch : BOOL;
    RightLimitSwitch : BOOL;
    GripLimitSwitch : BOOL;
    ReleaseLimitSwitch : BOOL;
END_VAR
VAR_OUTPUT
    MoveDown : BOOL;
    MoveUp : BOOL;
    MoveLeft : BOOL;
    MoveRight : BOOL;
    ActivateGrip : BOOL;
    ActivateRelease : BOOL;
END_VAR
VAR
    startTrig : R_TRIG;
    sdStep : INT := 0;
    autoStep : INT := 0;
    sdDone : BOOL;
    autoDone : BOOL;
    tmpMoveDown : BOOL;
    tmpMoveUp : BOOL;
    tmpMoveLeft : BOOL;
    tmpMoveRight : BOOL;
    tmpActivateGrip : BOOL;
    tmpActivateRelease : BOOL;
END_VAR

startTrig(CLK := Start);

tmpMoveDown := FALSE;
tmpMoveUp := FALSE;
tmpMoveLeft := FALSE;
tmpMoveRight := FALSE;
tmpActivateGrip := FALSE;
tmpActivateRelease := FALSE;

IF ManualMode THEN
    tmpMoveDown := DownButton AND NOT DownLimitSwitch;
    tmpMoveUp := UpButton AND NOT UpLimitSwitch;
    tmpMoveLeft := LeftButton AND NOT LeftLimitSwitch;
    tmpMoveRight := RightButton AND NOT RightLimitSwitch;
    tmpActivateGrip := GripButton AND NOT GripLimitSwitch;
    tmpActivateRelease := ReleaseButton AND NOT ReleaseLimitSwitch;

    IF tmpMoveDown AND tmpMoveUp THEN
        tmpMoveDown := FALSE;
        tmpMoveUp := FALSE;
    END_IF;
    IF tmpMoveLeft AND tmpMoveRight THEN
        tmpMoveLeft := FALSE;
        tmpMoveRight := FALSE;
    END_IF;
    IF tmpActivateGrip AND tmpActivateRelease THEN
        tmpActivateGrip := FALSE;
        tmpActivateRelease := FALSE;
    END_IF;

ELSIF SingleStepMode THEN
    CASE sdStep OF
        1: sdDone := DownLimitSwitch;
        2: sdDone := GripLimitSwitch;
        3: sdDone := UpLimitSwitch;
        4: sdDone := RightLimitSwitch;
        5: sdDone := DownLimitSwitch;
        6: sdDone := ReleaseLimitSwitch;
        7: sdDone := UpLimitSwitch;
        8: sdDone := LeftLimitSwitch;
    ELSE
        sdDone := TRUE;
    END_CASE;

    IF EmergencyStop AND startTrig.Q AND sdDone THEN
        IF sdStep >= 8 THEN
            sdStep := 1;
        ELSE
            sdStep := sdStep + 1;
        END_IF;
    END_IF;

    CASE sdStep OF
        1: tmpMoveDown := NOT DownLimitSwitch;
        2: tmpActivateGrip := NOT GripLimitSwitch;
        3: tmpMoveUp := NOT UpLimitSwitch;
        4: tmpMoveRight := NOT RightLimitSwitch;
        5: tmpMoveDown := NOT DownLimitSwitch;
        6: tmpActivateRelease := NOT ReleaseLimitSwitch;
        7: tmpMoveUp := NOT UpLimitSwitch;
        8: tmpMoveLeft := NOT LeftLimitSwitch;
    END_CASE;

ELSIF (SingleCycleMode OR ContinuousMode) THEN
    IF EmergencyStop AND startTrig.Q AND (autoStep = 0) THEN
        autoStep := 1;
    END_IF;

    CASE autoStep OF
        1: autoDone := DownLimitSwitch;
        2: autoDone := GripLimitSwitch;
        3: autoDone := UpLimitSwitch;
        4: autoDone := RightLimitSwitch;
        5: autoDone := DownLimitSwitch;
        6: autoDone := ReleaseLimitSwitch;
        7: autoDone := UpLimitSwitch;
        8: autoDone := LeftLimitSwitch;
    ELSE
        autoDone := TRUE;
    END_CASE;

    IF EmergencyStop AND (autoStep <> 0) AND autoDone THEN
        IF SingleCycleMode THEN
            IF autoStep < 8 THEN
                autoStep := autoStep + 1;
            ELSE
                autoStep := 0;
            END_IF;
        ELSIF ContinuousMode THEN
            IF autoStep < 8 THEN
                autoStep := autoStep + 1;
            ELSE
                autoStep := 1;
            END_IF;
        END_IF;
    END_IF;

    CASE autoStep OF
        1: tmpMoveDown := NOT DownLimitSwitch;
        2: tmpActivateGrip := NOT GripLimitSwitch;
        3: tmpMoveUp := NOT UpLimitSwitch;
        4: tmpMoveRight := NOT RightLimitSwitch;
        5: tmpMoveDown := NOT DownLimitSwitch;
        6: tmpActivateRelease := NOT ReleaseLimitSwitch;
        7: tmpMoveUp := NOT UpLimitSwitch;
        8: tmpMoveLeft := NOT LeftLimitSwitch;
    END_CASE;

END_IF;

IF NOT EmergencyStop THEN
    MoveDown := FALSE;
    MoveUp := FALSE;
    MoveLeft := FALSE;
    MoveRight := FALSE;
    ActivateGrip := FALSE;
    ActivateRelease := FALSE;
ELSE
    MoveDown := tmpMoveDown;
    MoveUp := tmpMoveUp;
    MoveLeft := tmpMoveLeft;
    MoveRight := tmpMoveRight;
    ActivateGrip := tmpActivateGrip;
    ActivateRelease := tmpActivateRelease;
END_IF;

END_FUNCTION_BLOCK

(* ---- public-medium-04.candidate_01.st ---- *)
FUNCTION_BLOCK FB_TemperatureControl
VAR_INPUT
    TemperatureSensorInput : REAL;
    SetTemperature : REAL;
END_VAR
VAR_OUTPUT
    CurrentTemperature : REAL;
    SetTempDisplay : REAL;
    HeaterStatus : BOOL;
    OverheatProtection : BOOL;
    HeaterOutput : BOOL;
END_VAR
VAR
    tmp_sensor_fault : BOOL;
    tmp_heat_allowed : BOOL;
    tmp_overheat_active : BOOL;
    tmp_heat_on_timer : TON;
    tmp_cooldown_timer : TON;
    tmp_heat_limit : TIME := T#5001MS;  (* strictly > 5 s continuous heating *)
    tmp_cooldown_limit : TIME := T#3S;
END_VAR

(*
ENGINEERING_CONTRACT
- CurrentTemperature/SetTempDisplay: combinational echoes, raw units.
- HeaterOutput: on when sensor valid, no overheat, sensor < set;
  off when sensor >= set, sensor fault, or overheat. Equal is off.
- OverheatProtection: latched TRUE on continuous heater on >5s; auto clear after 3s cooldown.
- HeaterStatus: echo of HeaterOutput.
- Sensor fault: <0.0 or >100.0. Fault and overheat force heater off.
- Unspecified: equal setpoint and reset after cooldown interpreted as above.
- PUB001-PUB008.
*)

(* CONTRACT_RULES [] *)

tmp_sensor_fault := (TemperatureSensorInput < 0.0) OR (TemperatureSensorInput > 100.0);

tmp_heat_allowed := (NOT tmp_sensor_fault)
                    AND (NOT tmp_overheat_active)
                    AND (TemperatureSensorInput < SetTemperature);

tmp_heat_on_timer(IN := tmp_heat_allowed, PT := tmp_heat_limit);

IF tmp_heat_on_timer.Q THEN
    tmp_overheat_active := TRUE;
END_IF;

tmp_cooldown_timer(IN := tmp_overheat_active, PT := tmp_cooldown_limit);

IF tmp_cooldown_timer.Q THEN
    tmp_overheat_active := FALSE;
    tmp_heat_allowed := (NOT tmp_sensor_fault)
                        AND (NOT tmp_overheat_active)
                        AND (TemperatureSensorInput < SetTemperature);
    tmp_heat_on_timer(IN := tmp_heat_allowed, PT := tmp_heat_limit);
END_IF;

HeaterOutput := (NOT tmp_sensor_fault)
                AND (NOT tmp_overheat_active)
                AND (TemperatureSensorInput < SetTemperature);

HeaterStatus := HeaterOutput;
OverheatProtection := tmp_overheat_active;
CurrentTemperature := TemperatureSensorInput;
SetTempDisplay := SetTemperature;

END_FUNCTION_BLOCK

(* ---- public-medium-04.patch_base_01.st ---- *)
FUNCTION_BLOCK FB_TemperatureControl
VAR_INPUT
    TemperatureSensorInput : REAL;
    SetTemperature : REAL;
END_VAR
VAR_OUTPUT
    CurrentTemperature : REAL;
    SetTempDisplay : REAL;
    HeaterStatus : BOOL;
    OverheatProtection : BOOL;
    HeaterOutput : BOOL;
END_VAR
VAR
    tmp_sensor_fault : BOOL;
    tmp_heat_allowed : BOOL;
    tmp_overheat_active : BOOL;
    tmp_heat_on_timer : TON;
    tmp_cooldown_timer : TON;
    tmp_heat_limit : TIME := T#5001MS;  (* strictly > 5 s continuous heating *)
    tmp_cooldown_limit : TIME := T#3S;
END_VAR

(*
ENGINEERING_CONTRACT
- CurrentTemperature/SetTempDisplay: combinational echoes, raw units.
- HeaterOutput: on when sensor valid, no overheat, sensor < set;
  off when sensor >= set, sensor fault, or overheat. Equal is off.
- OverheatProtection: latched TRUE on continuous heater on >5s; auto clear after 3s cooldown.
- HeaterStatus: echo of HeaterOutput.
- Sensor fault: <0.0 or >100.0. Fault and overheat force heater off.
- Unspecified: equal setpoint and reset after cooldown interpreted as above.
- PUB001-PUB008.
*)

(* CONTRACT_RULES [] *)

tmp_sensor_fault := (TemperatureSensorInput < 0.0) OR (TemperatureSensorInput > 100.0);

tmp_heat_allowed := (NOT tmp_sensor_fault)
                    AND (NOT tmp_overheat_active)
                    AND (TemperatureSensorInput < SetTemperature);

tmp_heat_on_timer(IN := tmp_heat_allowed, PT := tmp_heat_limit);

IF tmp_heat_on_timer.Q THEN
    tmp_overheat_active := TRUE;
END_IF;

tmp_cooldown_timer(IN := tmp_overheat_active, PT := tmp_cooldown_limit);

IF tmp_cooldown_timer.Q THEN
    tmp_overheat_active := FALSE;
END_IF;

HeaterOutput := (NOT tmp_sensor_fault)
                AND (NOT tmp_overheat_active)
                AND (TemperatureSensorInput < SetTemperature);

HeaterStatus := HeaterOutput;
OverheatProtection := tmp_overheat_active;
CurrentTemperature := TemperatureSensorInput;
SetTempDisplay := SetTemperature;

END_FUNCTION_BLOCK

(* ---- public-medium-04.raw_candidate_01.st ---- *)
FUNCTION_BLOCK FB_TemperatureControl
VAR_INPUT
    TemperatureSensorInput : REAL;
    SetTemperature : REAL;
END_VAR
VAR_OUTPUT
    CurrentTemperature : REAL;
    SetTempDisplay : REAL;
    HeaterStatus : BOOL;
    OverheatProtection : BOOL;
    HeaterOutput : BOOL;
END_VAR
VAR
    tmp_sensor_fault : BOOL;
    tmp_heat_allowed : BOOL;
    tmp_overheat_active : BOOL;
    tmp_heat_on_timer : TON;
    tmp_cooldown_timer : TON;
    tmp_heat_limit : TIME := T#5001MS;  (* strictly > 5 s continuous heating *)
    tmp_cooldown_limit : TIME := T#3S;
END_VAR

(*
ENGINEERING_CONTRACT
- CurrentTemperature/SetTempDisplay: combinational echoes, raw units.
- HeaterOutput: on when sensor valid, no overheat, sensor < set;
  off when sensor >= set, sensor fault, or overheat. Equal is off.
- OverheatProtection: latched TRUE on continuous heater on >5s; auto clear after 3s cooldown.
- HeaterStatus: echo of HeaterOutput.
- Sensor fault: <0.0 or >100.0. Fault and overheat force heater off.
- Unspecified: equal setpoint and reset after cooldown interpreted as above.
- PUB001-PUB008.
*)

(* CONTRACT_RULES [] *)

tmp_sensor_fault := (TemperatureSensorInput < 0.0) OR (TemperatureSensorInput > 100.0);

tmp_heat_allowed := (NOT tmp_sensor_fault)
                    AND (NOT tmp_overheat_active)
                    AND (TemperatureSensorInput < SetTemperature);

tmp_heat_on_timer(IN := tmp_heat_allowed, PT := tmp_heat_limit);

IF tmp_heat_on_timer.Q THEN
    tmp_overheat_active := TRUE;
END_IF;

tmp_cooldown_timer(IN := tmp_overheat_active, PT := tmp_cooldown_limit);

IF tmp_cooldown_timer.Q THEN
    tmp_overheat_active := FALSE;
    tmp_heat_allowed := (NOT tmp_sensor_fault)
                        AND (NOT tmp_overheat_active)
                        AND (TemperatureSensorInput < SetTemperature);
    tmp_heat_on_timer(IN := tmp_heat_allowed, PT := tmp_heat_limit);
END_IF;

HeaterOutput := (NOT tmp_sensor_fault)
                AND (NOT tmp_overheat_active)
                AND (TemperatureSensorInput < SetTemperature);

HeaterStatus := HeaterOutput;
OverheatProtection := tmp_overheat_active;
CurrentTemperature := TemperatureSensorInput;
SetTempDisplay := SetTemperature;

END_FUNCTION_BLOCK
